(* IEC 61131-3 sources: labSCADA/project-view, 13 files *)

(* ---- FB_AnalogAlarm.st ---- *)
(* ==============================================================================
   FUNCTION BLOCK: FB_AnalogAlarm
   DESCRIPTION: IEC 61131-3 Structured Text implementation of an SEL RTAC-style
                analog alarm monitor with pickup/dropout hysteresis deadbands
                and sustained excursion / reset timers.

                Supports:
                - High Alarm trip / dropout (e.g. Fridge High > 8.0°C, reset < 7.5°C)
                - Low Alarm trip / dropout (e.g. Fridge Low < 2.0°C, reset > 2.5°C)
                - Window Alarm (High + Low simultaneously enabled)
                - Configurable Pickup Delay (prevents trips on brief door opens or noise)
                - Configurable Dropout Delay (anti-chatter filter on recovery)
                - Diagnostic Trip Outputs (HighTrip, LowTrip, Elapsed Timers)
   ============================================================================== *)
FUNCTION_BLOCK FB_AnalogAlarm
VAR_INPUT
	rVal            : REAL;             (* Analog process value to monitor (e.g. Temperature) *)
    bEnableHigh     : BOOL := TRUE;     (* Enable High Alarm monitoring *)
    rHighPickup     : REAL := 0.0;      (* High trip pickup threshold *)
    rHighDropout    : REAL := 0.0;      (* High trip reset threshold (or leave 0.0 and use rHysteresis) *)
    bEnableLow      : BOOL := FALSE;    (* Enable Low Alarm monitoring *)
    rLowPickup      : REAL := 0.0;      (* Low trip pickup threshold *)
    rLowDropout     : REAL := 0.0;      (* Low trip reset threshold (or leave 0.0 and use rHysteresis) *)
    rHysteresis     : REAL := 0.0;      (* Optional deadband offset applied if Dropout not explicitly set *)
    tPickupDelay    : TIME := T#0S;     (* Time excursion must persist before alarm asserts *)
    tDropoutDelay   : TIME := T#0S;     (* Time normal state must persist before alarm clears *)
END_VAR
VAR_OUTPUT
	bAlarm          : BOOL := FALSE;    (* Filtered alarm output (Active Alarm) *)
    bWarn           : BOOL := FALSE;    (* Pre-alarm warning: In excursion (pickup), timing towards alarm *)
    bPickup         : BOOL := FALSE;    (* Instantaneous pickup status (pre-timer) *)
    bHighTrip       : BOOL := FALSE;    (* TRUE if High Alarm condition caused/maintains trip *)
    bLowTrip        : BOOL := FALSE;    (* TRUE if Low Alarm condition caused/maintains trip *)
    tElapsedPU      : TIME := T#0S;     (* Current elapsed pickup timer *)
    tElapsedDO      : TIME := T#0S;     (* Current elapsed dropout timer *)
END_VAR
VAR
	rEffHighDO      : REAL;
    rEffLowDO       : REAL;
    bHighCondition  : BOOL := FALSE;
    bLowCondition   : BOOL := FALSE;
    fbTimer         : FB_PickupDropout;
END_VAR
// --- implementation ---
// 1. Calculate effective dropout thresholds
IF rHighDropout <> 0.0 THEN
    rEffHighDO := rHighDropout;
ELSIF rHysteresis > 0.0 THEN
    rEffHighDO := rHighPickup - rHysteresis;
ELSE
    rEffHighDO := rHighPickup;
END_IF;

IF rLowDropout <> 0.0 THEN
    rEffLowDO := rLowDropout;
ELSIF rHysteresis > 0.0 THEN
    rEffLowDO := rLowPickup + rHysteresis;
ELSE
    rEffLowDO := rLowPickup;
END_IF;

// 2. High threshold hysteresis evaluation
IF bEnableHigh THEN
    IF rVal >= rHighPickup THEN
        bHighCondition := TRUE;
    ELSIF rVal <= rEffHighDO THEN
        bHighCondition := FALSE;
    END_IF;
ELSE
    bHighCondition := FALSE;
END_IF;

// 3. Low threshold hysteresis evaluation
IF bEnableLow THEN
    IF rVal <= rLowPickup THEN
        bLowCondition := TRUE;
    ELSIF rVal >= rEffLowDO THEN
        bLowCondition := FALSE;
    END_IF;
ELSE
    bLowCondition := FALSE;
END_IF;

// 4. Pickup / Dropout timing filter (SEL RTAC PU_DO equivalent)
fbTimer(
    IN := (bHighCondition OR bLowCondition),
    tPickupDelay := tPickupDelay,
    tDropoutDelay := tDropoutDelay
);

bAlarm     := fbTimer.Q;
bPickup    := fbTimer.bPickup;
bWarn      := fbTimer.bPickup AND NOT fbTimer.Q;
tElapsedPU := fbTimer.tElapsedPU;
tElapsedDO := fbTimer.tElapsedDO;

// 5. Diagnostic cause flags
IF bAlarm THEN
    bHighTrip := bHighCondition;
    bLowTrip  := bLowCondition;
ELSE
    bHighTrip := FALSE;
    bLowTrip  := FALSE;
END_IF;
END_FUNCTION

(* ---- FB_APC_SmartUPS.st ---- *)
(* ==============================================================================
   FUNCTION BLOCK: FB_APC_SmartUPS
   DESCRIPTION: Encapsulated clinical monitoring block for UPS Power Systems
                following the Schneider Electric / APC Smart-UPS Modbus Register Map
                (AN-176 / 990-9840).
                - Supervised Utility Grid Power Loss (Generator Dispatch)
                - Battery State of Charge & Remaining Runtime Monitoring
                - Low Battery Reserve Emergency Escalation
                - Beeper Mute / Silence Supervisory Command Control
   ============================================================================== *)
FUNCTION_BLOCK FB_APC_SmartUPS
VAR_INPUT
    wStatusWord         : WORD := 16#0001;  (* Register 40001: Bit 0=Online, Bit 1=On Battery, Bit 4=Low Battery *)
    wBatteryPct         : WORD := 100;     (* Register 40002: Battery Charge (0-100%) *)
    wRuntimeSec         : WORD := 0;       (* Register 40003: Runtime in seconds *)
    wLineVoltageX10     : WORD := 1200;    (* Register 40004: Line Voltage * 10 (1200 = 120.0 V) *)
    wLoadPct            : WORD := 0;       (* Register 40005: Inverter Load (0-100%) *)
    wRuntimeMin         : WORD := 60;      (* Register 40007: Runtime in minutes *)
    wBeeperStatus       : WORD := 1;       (* Register 40008: 1=Enabled, 2=Muted, 3=Disabled *)

    (* --- Interactive Operator Commands (from Kiosk UI or PLC) --- *)
    bCmdMuteBeeper      : BOOL := FALSE;   (* TRUE pulse: Temporarily mute beeper for current power loss *)
    bCmdDisableBeeper   : BOOL := FALSE;   (* TRUE pulse: Disable beeper speaker *)
    bCmdEnableBeeper    : BOOL := FALSE;   (* TRUE pulse: Enable beeper speaker *)

    tPowerLossDelay     : TIME := T#10S;   (* Debounce filter to ignore momentary utility grid flickers *)
    wLowBatteryLimit    : WORD := 20;      (* Low battery alarm threshold (%) *)
    wLowRuntimeLimitMin : WORD := 15;      (* Low runtime alarm threshold (minutes) *)
END_VAR
VAR_OUTPUT
    bOnline             : BOOL := TRUE;    (* TRUE = Grid utility power is normal *)
    bOnBattery          : BOOL := FALSE;   (* TRUE = Running on battery inverter *)
    bAlarmPowerLost     : BOOL := FALSE;   (* Priority 2: Utility grid dropped -> Manual generator required *)
    bAlarmLowBattery    : BOOL := FALSE;   (* Priority 1: Battery reserve critically low *)
    rBatteryPct         : REAL := 100.0;   (* Battery % (0.0 - 100.0) *)
    rLineVoltage        : REAL := 120.0;   (* Utility line voltage in Volts RMS *)
    rRuntimeMinutes     : REAL := 60.0;    (* Estimated remaining runtime in minutes *)
    rLoadPct            : REAL := 0.0;     (* Current load percentage *)
    bBeeperMuted        : BOOL := FALSE;   (* Beeper is currently muted *)
    bBeeperDisabled     : BOOL := FALSE;   (* Beeper is disabled *)

    (* --- Modbus Command Output (Mapped to Holding Register 40010 / Offset 9) --- *)
    wCommandOut         : WORD := 0;       (* 1=Mute, 2=Disable, 3=Enable *)
END_VAR
VAR
    fbFilterPowerLoss   : FB_PickupDropout;
    tonCmdPulse         : TON;
    wActiveCmd          : WORD := 0;
    bPrevMute           : BOOL := FALSE;
    bPrevDisable        : BOOL := FALSE;
    bPrevEnable         : BOOL := FALSE;
END_VAR
// --- implementation ---
// 1. DECODE APC SMART-UPS STATUS WORD (Register 40001)
// Bit 0 = State Online (Grid OK)
// Bit 1 = State On Battery (Power Failure)
// Bit 4 = Low Battery
bOnline    := (wStatusWord AND 16#0001) <> 0;
bOnBattery := (wStatusWord AND 16#0002) <> 0;

// 2. CONVERT RAW TELEMETRY TO ENGINEERING UNITS
rBatteryPct     := WORD_TO_REAL(wBatteryPct);
rLineVoltage    := WORD_TO_REAL(wLineVoltageX10) / 10.0;
rLoadPct        := WORD_TO_REAL(wLoadPct);

// Beeper status
bBeeperMuted    := (wBeeperStatus = 2);
bBeeperDisabled := (wBeeperStatus = 3);

// Calculate runtime in minutes (prefer wRuntimeMin if non-zero, else wRuntimeSec / 60)
IF wRuntimeMin > 0 THEN
    rRuntimeMinutes := WORD_TO_REAL(wRuntimeMin);
ELSIF wRuntimeSec > 0 THEN
    rRuntimeMinutes := WORD_TO_REAL(wRuntimeSec) / 60.0;
ELSE
    rRuntimeMinutes := 0.0;
END_IF;

// 3. DEBOUNCED UTILITY POWER LOSS ALARM (Generator Dispatch)
// Ignores 1-2 second lightning flickers, trips after sustained outage (tPowerLossDelay)
fbFilterPowerLoss(
    IN            := bOnBattery,
    tPickupDelay  := tPowerLossDelay,
    tDropoutDelay := T#5S
);
bAlarmPowerLost := fbFilterPowerLoss.Q;

// 4. CRITICAL LOW BATTERY ALARM
// Triggers if battery % drops below limit OR runtime drops below critical threshold while on battery
IF bOnBattery AND ((wBatteryPct <= wLowBatteryLimit) OR (rRuntimeMinutes <= WORD_TO_REAL(wLowRuntimeLimitMin))) THEN
    bAlarmLowBattery := TRUE;
ELSE
    bAlarmLowBattery := FALSE;
END_IF;

// 5. BEEPER COMMAND EXECUTION (Pulsed Output to Modbus Register 40010)
// Latch active command for 1.5s so asynchronous Modbus cyclic task reliably transmits write
IF bCmdMuteBeeper AND NOT bPrevMute THEN
    wActiveCmd := 1;       // 1 = Mute
    bCmdMuteBeeper := FALSE;
ELSIF bCmdDisableBeeper AND NOT bPrevDisable THEN
    wActiveCmd := 2;       // 2 = Disable
    bCmdDisableBeeper := FALSE;
ELSIF bCmdEnableBeeper AND NOT bPrevEnable THEN
    wActiveCmd := 3;       // 3 = Enable
    bCmdEnableBeeper := FALSE;
END_IF;

bPrevMute    := bCmdMuteBeeper;
bPrevDisable := bCmdDisableBeeper;
bPrevEnable  := bCmdEnableBeeper;

tonCmdPulse(IN := (wActiveCmd > 0), PT := T#1500MS);
IF tonCmdPulse.Q THEN
    wActiveCmd := 0;
END_IF;

wCommandOut := wActiveCmd;
END_FUNCTION

(* ---- FB_Dewar.st ---- *)
(* ==============================================================================
   FUNCTION BLOCK: FB_Dewar
   DESCRIPTION: Encapsulated clinical monitoring block for Liquid Nitrogen (LN2)
                cryogenic storage vessels (dewars / freezers).
                - Scaled raw integer input (iRawTempX10 / 10.0 -> °C)
                - High threshold alarm with hysteresis & debounced pickup timing
                - Clinical fault supervision (Open circuit, wiring short, comms loss)
                - High-temperature excursion alarm gated off during hardware faults
                - Wireless cleanroom health diagnostics (Battery, RSSI, Watchdog, Faults)
   ============================================================================== *)
FUNCTION_BLOCK FB_Dewar
VAR_INPUT
    (* --- Operational Alarm Thresholds & Delays --- *)
    rHighTrip           : REAL := -135.0;   (* Critical specimen danger limit (°C) *)
    rHysteresis         : REAL := 5.0;      (* Reset deadband (°C) *)
    tPickupDelay        : TIME := T#30S;    (* Sustained warm excursion required to trip *)
    tDropoutDelay       : TIME := T#10S;    (* Clean fill required to reset *)

    (* --- 8 Modbus Holding Registers (Direct from Bridge Slot 1) --- *)
    wRawTempX10         : WORD := 16#D8F0;  (* Offset 0: Dewar scaled temp * 10 (-1954 = -195.4 °C, -9999 = Sentinel) *)
    uiRawBatteryMv      : UINT := 3850;     (* Offset 1: Battery health in millivolts *)
    uiRawFaultCode      : UINT := 0;        (* Offset 2: Probe fault (0=OK, 1=Open, 2=GND, 3=VCC, 4=Hardware Error) *)
    wRawRSSI            : WORD := 16#FFCE;  (* Offset 3: Wireless link margin in dBm (-50 = 16#FFCE) *)
    wRawSeqLow          : WORD := 0;        (* Offset 4: Sequence counter low word *)
    wRawSeqHigh         : WORD := 0;        (* Offset 5: Sequence counter high word *)
    uiRawAgeSec         : UINT := 0;        (* Offset 6: Telemetry age in seconds *)
    wRawStatusFlags     : WORD := 16#0001;  (* Offset 7: Bit 0=Online, Bit 1=LowBatt, Bit 2=CommLoss, Bit 3=AccessMode *)
    bIsWireless         : BOOL := TRUE;     (* TRUE = Enable wireless diagnostics *)
    tCommLossTimeout    : TIME := T#60S;    (* Watchdog comms loss alarm threshold *)

    (* --- Interactive Operator Commands (from Kiosk UI or OPC UA) --- *)
    bCmdSetAccessMode   : BOOL := FALSE;    (* TRUE pulse: Activate Access Mode (Alarms paused 30 min) *)
    bCmdCancelAccessMode: BOOL := FALSE;    (* TRUE pulse: Cancel Access Mode immediately *)
    rCalOffset          : REAL := 0.0;      (* NIST calibration trim offset in °C (clamped +/-10.0) *)
END_VAR
VAR_OUTPUT
    rProcessTemp        : REAL := -999.0;   (* Published process temperature to SCADA (°C) *)
    bAlarm              : BOOL := FALSE;    (* Priority 2 Emergency Temperature Alarm flag *)
    bWarn               : BOOL := FALSE;    (* Pre-alarm pickup delay warning flag *)
    rBatteryVolts       : REAL := 3.85;     (* Published battery voltage (V) *)
    bLowBattery         : BOOL := FALSE;    (* Low battery warning flag (< 3.4V) *)
    iRSSI               : INT := -50;       (* Published wireless link margin (dBm) *)
    bCommLoss           : BOOL := FALSE;    (* Comms loss watchdog alarm *)
    bProbeFault         : BOOL := TRUE;     (* Physical probe disconnected or shorted (defaults TRUE on cold boot) *)
    uiFaultCode         : UINT := 0;        (* Published probe fault reason (0=OK, 1=Open, 2=GND, 3=VCC) *)
    uiAgeSec            : UINT := 0;        (* Telemetry age in seconds *)
    bAccessMode         : BOOL := FALSE;    (* Access Mode active - Alarms paused 30 min for tank maintenance *)

    (* --- Modbus Command Outputs (Mapped to Bridge Holding Regs 10 & 11) --- *)
    wCommandMailboxOut  : WORD := 0;        (* Offset 10: 5 = SetAccessMode *)
    wCommandParamOut    : WORD := 0;        (* Offset 11: 30 = 30 minutes, 0 = Cancel *)
END_VAR
VAR
    iTempX10            : INT;
    fbAlarmEval         : FB_AnalogAlarm;
    wActiveCmdCode      : WORD := 0;
    wActiveCmdParam     : WORD := 0;
    bPrevSetAccess      : BOOL := FALSE;
    bPrevCancelAccess   : BOOL := FALSE;
    tonCmdPulse         : TON;
    rCalOffsetEff       : REAL := 0.0;
END_VAR
VAR CONSTANT
    cMaxCalOffset       : REAL := 10.0;
END_VAR
// --- implementation ---
// ==============================================================================
// 1. HARDWARE HEALTH & TELEMETRY DECODING
// ==============================================================================
// Explicitly cast Modbus unsigned WORD inputs to signed two's complement INT
iTempX10 := TO_INT(wRawTempX10);

IF bIsWireless THEN
    rBatteryVolts := TO_REAL(uiRawBatteryMv) / 1000.0;
    bLowBattery   := (uiRawBatteryMv < 3400) OR (wRawStatusFlags.1);
    iRSSI         := TO_INT(wRawRSSI);
    uiAgeSec      := uiRawAgeSec;
    uiFaultCode   := uiRawFaultCode;

    // Probe fault if hardware reported fault code or value is sentinel (<= -273°C or >= 900°C)
    bProbeFault   := (uiRawFaultCode <> 0) OR (iTempX10 <= -2730) OR (iTempX10 >= 9000);

    // Watchdog comms loss if bridge flagged or age exceeds timeout
    bCommLoss     := (NOT wRawStatusFlags.0) OR (wRawStatusFlags.2) OR (uiRawAgeSec > (TIME_TO_UINT(tCommLossTimeout) / 1000));

    // Access Mode Active (Bit 3 of status flags: Alarms paused 30 min)
    bAccessMode   := wRawStatusFlags.3;
ELSE
    rBatteryVolts := 0.0;
    bLowBattery   := FALSE;
    iRSSI         := 0;
    bCommLoss     := FALSE;
    uiFaultCode   := 0;
    bProbeFault   := (iTempX10 <= -2730) OR (iTempX10 >= 9000);
    uiAgeSec      := 0;
    bAccessMode   := FALSE;
END_IF;

// ==============================================================================
// 2. TEMPERATURE SENTINEL MAPPING
// ==============================================================================
IF rCalOffset > cMaxCalOffset THEN
    rCalOffsetEff := cMaxCalOffset;
ELSIF rCalOffset < -cMaxCalOffset THEN
    rCalOffsetEff := -cMaxCalOffset;
ELSE
    rCalOffsetEff := rCalOffset;
END_IF;

// If probe is faulted or comms lost, output standard invalid sentinel (-999.0 °C)
IF bProbeFault OR bCommLoss THEN
    rProcessTemp := -999.0;
ELSE
    rProcessTemp := (TO_REAL(iTempX10) / 10.0) + rCalOffsetEff;
END_IF;

// ==============================================================================
// 3. CLINICAL ALARM EVALUATION (Pickup / Dropout & Hysteresis)
// ==============================================================================
// Thermal excursion alarms are only evaluated when sensor data is valid and not in access mode
fbAlarmEval(
    rVal          := rProcessTemp,
    bEnableHigh   := NOT (bProbeFault OR bCommLoss OR bAccessMode),
    rHighPickup   := rHighTrip,
    rHighDropout  := rHighTrip - rHysteresis,
    bEnableLow    := FALSE,
    tPickupDelay  := tPickupDelay,
    tDropoutDelay := tDropoutDelay
);

// If in Access Mode, clamp alarms and warnings to FALSE immediately (bypassing dropout timer)
IF bAccessMode THEN
    bAlarm := FALSE;
    bWarn  := FALSE;
ELSE
    bAlarm := fbAlarmEval.bAlarm;
    bWarn  := fbAlarmEval.bWarn;
END_IF;

// ==============================================================================
// 4. SUPERVISORY COMMAND DISPATCH (Downlink to Bridge & Physical Node)
// ==============================================================================
// Latch active command for 2.0s so Modbus cyclic write task reliably transmits to Bridge
IF bCmdSetAccessMode AND NOT bPrevSetAccess THEN
    wActiveCmdCode    := 5;     // 5 = SetAccessMode
    wActiveCmdParam   := 30;    // 30 minutes
    bCmdSetAccessMode := FALSE;
ELSIF bCmdCancelAccessMode AND NOT bPrevCancelAccess THEN
    wActiveCmdCode       := 5;  // 5 = SetAccessMode
    wActiveCmdParam      := 0;  // 0 = Cancel / Normal Mode
    bCmdCancelAccessMode := FALSE;
END_IF;

bPrevSetAccess    := bCmdSetAccessMode;
bPrevCancelAccess := bCmdCancelAccessMode;

tonCmdPulse(IN := (wActiveCmdCode > 0), PT := T#2000MS);
IF tonCmdPulse.Q THEN
    wActiveCmdCode  := 0;
    wActiveCmdParam := 0;
END_IF;

wCommandMailboxOut := wActiveCmdCode;
wCommandParamOut   := wActiveCmdParam;
END_FUNCTION

(* ---- FB_FacilityDoor.st ---- *)
(* ==============================================================================
   FUNCTION BLOCK: FB_FacilityDoor
   DESCRIPTION: Encapsulated monitoring block for cleanroom and facility access doors
                (Main Entry, Procedure Room, Cryo Storage, Air Shower, Gown In/Out).
                Features:
                - Fail-safe normally closed contact supervision (24V/TRUE = Closed, 0V/FALSE = Open / Unwired)
                - Sustained open timer with contact chatter dropout filter (FB_PickupDropout)
                - Direct physical terminal binding (bDoorClosed)
                - Filtered alarm output to SCADA (bDoorAlarm)
   ============================================================================== *)
FUNCTION_BLOCK FB_FacilityDoor
VAR_INPUT
    bDoorClosed         : BOOL := FALSE;    (* Hardware DI: 24V/TRUE = Closed, 0V/FALSE = Open / Unwired *)
    tOpenAlarmDelay     : TIME := T#60M;    (* Sustained open threshold before alarm asserts *)
    tDropoutDelay       : TIME := T#5S;     (* Anti-chatter filter on door closure *)
END_VAR
VAR_OUTPUT
    bDoorAlarm          : BOOL := FALSE;    (* Filtered Priority 2 Alarm output to SCADA *)
END_VAR
VAR
    fbFilter            : FB_PickupDropout;
END_VAR
// --- implementation ---
// TIMED DEBOUNCE FILTER FOR DOOR HELD OPEN ALARM
fbFilter(
    IN            := NOT bDoorClosed,
    tPickupDelay  := tOpenAlarmDelay,
    tDropoutDelay := tDropoutDelay
);
bDoorAlarm := fbFilter.Q;
END_FUNCTION

(* ---- FB_G210_Incubator.st ---- *)
(* ==============================================================================
   FUNCTION BLOCK: FB_G210_Incubator
   DESCRIPTION: Encapsulated clinical monitoring block for K-Systems G210
                Multi-Chamber Incubators (10 Heated Zones).
                - 10 Chamber Zone Temperatures (Default -99.0°C unassigned sentinel)
                - Direct Physical Dry Alarm Contact (bAlarmContact)
                - Door/Recovery Mute Supervision (bMute)
                - Pickup/Dropout Debounce Filter
   ============================================================================== *)
FUNCTION_BLOCK FB_G210_Incubator
VAR_INPUT
    bAlarmContact       : BOOL := FALSE;    (* Physical dry alarm contact from incubator (Fail-Safe NC: TRUE = Normal/Closed, FALSE = Alarm/Open) *)
    bMute               : BOOL := FALSE;    (* TRUE = Suppress alarm (Cabinet door open or recovery grace) *)
    tPickupDelay        : TIME := T#15S;    (* Contact bounce filter *)
    tDropoutDelay       : TIME := T#5S;     (* Recovery confirmation filter *)
END_VAR
VAR_OUTPUT
    bAlarm              : BOOL := FALSE;    (* Filtered Priority 2 Alarm output to SCADA *)
    bMuted              : BOOL := FALSE;    (* Contact is tripped but actively suppressed by cabinet mute *)
    rZoneTemps          : ARRAY[1..10] OF REAL := [10(-99.0)];  (* 10 Heated Chambers, Default -99.0 °C (Unwired Sentinel) *)
END_VAR
VAR
    fbFilter            : FB_PickupDropout;
END_VAR
// --- implementation ---
// 1. TIMED DEBOUNCE FILTER ON FAIL-SAFE NC ALARM CONTACT (TRUE = Closed/Normal, FALSE = Open/Alarm)
fbFilter(
    IN            := NOT bAlarmContact,
    tPickupDelay  := tPickupDelay,
    tDropoutDelay := tDropoutDelay
);

// 2. MUTE SUPERVISION
// When bMute is TRUE (cabinet door open or grace period), suppress bAlarm.
bMuted := bMute AND fbFilter.Q;

IF bMute THEN
    bAlarm := FALSE;
ELSE
    bAlarm := fbFilter.Q;
END_IF;
END_FUNCTION

(* ---- FB_Incubator.st ---- *)
(* ==============================================================================
   FUNCTION BLOCK: FB_Incubator
   DESCRIPTION: Encapsulated clinical monitoring block for Embryology Incubators
                (benchtop trigas, box incubators) via discrete dry alarm contacts.
                Features:
                - Pickup/Dropout debounce filter (FB_PickupDropout)
                - Direct physical terminal binding (bAlarmContact)
                - Cabinet door / post-close mute supervision (bMute)
   ============================================================================== *)
FUNCTION_BLOCK FB_Incubator
VAR_INPUT
    bAlarmContact       : BOOL := FALSE;    (* Physical dry alarm contact from incubator (FALSE = Normal, TRUE = Alarm) *)
    bMute               : BOOL := FALSE;    (* TRUE = Suppress alarm (Cabinet door open or recovery grace) *)
    tPickupDelay        : TIME := T#15S;    (* Contact bounce suppression filter *)
    tDropoutDelay       : TIME := T#5S;     (* Recovery confirmation filter *)
END_VAR
VAR_OUTPUT
    bAlarm              : BOOL := FALSE;    (* Filtered Priority 2 Alarm output to SCADA *)
    bMuted              : BOOL := FALSE;    (* Contact is tripped but suppressed by active mute *)
END_VAR
VAR
    fbFilter            : FB_PickupDropout;
END_VAR
// --- implementation ---
// 1. TIMED DEBOUNCE FILTER
fbFilter(
    IN            := bAlarmContact,
    tPickupDelay  := tPickupDelay,
    tDropoutDelay := tDropoutDelay
);

// 2. MUTE SUPERVISION
// When bMute is active (cabinet door open or post-close grace), suppress bAlarm.
bMuted := bMute AND fbFilter.Q;

IF bMute THEN
    bAlarm := FALSE;
ELSE
    bAlarm := fbFilter.Q;
END_IF;
END_FUNCTION

(* ---- FB_IncubatorCabinet.st ---- *)
(* ==============================================================================
   FUNCTION BLOCK: FB_IncubatorCabinet
   DESCRIPTION: Enclosure microclimate and access supervision for benchtop
                incubator cabinet.
                Features:
                - Standardized fail-safe door contact supervision (Closed loop = Closed, Open loop = Open)
                - Autonomous incubator alarm muting while door is open
                - Post-closure recovery grace timer (TOF) to prevent nuisance alarms
                - Cabinet door left open alarm (TON)
                - Thermostatic exhaust fan control loop (hysteresis)
   ============================================================================== *)
FUNCTION_BLOCK FB_IncubatorCabinet
VAR_INPUT
    bDoorClosed         : BOOL := FALSE;    (* Hardware DI: 24V/TRUE = Closed, 0V/FALSE = Open / Disconnected *)
    tDoorAlarmDelay     : TIME := T#3M;     (* Alarm if cabinet door left open longer than this *)
    tPostCloseGrace     : TIME := T#3M;     (* Time to keep incubator alarms muted after door closes *)
    wRawTempX10         : WORD := 16#D8F0;  (* Raw Modbus 750-461 register x10 (244 = 24.4°C, -9999 = 16#D8F0) *)
    rFanOnSetpoint      : REAL := 28.0;     (* Exhaust fan ON setpoint in °C *)
    rFanHysteresis      : REAL := 1.5;      (* Deadband in °C (turns off at 26.5°C) *)
    rCalOffset          : REAL := 0.0;      (* NIST calibration trim offset in °C (clamped +/-10.0) *)
END_VAR
VAR_OUTPUT
    bDoorAlarm          : BOOL := FALSE;    (* Alarm: Cabinet door held open past delay *)
    bIncubatorMute      : BOOL := FALSE;    (* TRUE while door is open OR during post-closure grace *)
    tGraceRemaining     : TIME := T#0S;     (* Time remaining in post-close recovery grace *)
    bFanCommand         : BOOL := FALSE;    (* Command to future DO fan relay *)
    bCabinetOvertemp    : BOOL := FALSE;    (* Alarm: Cabinet internal temp >= 32°C *)
    rProcessTemp        : REAL := -999.0;   (* Published cabinet temperature (°C) to SCADA & DB *)
    bProbeFault         : BOOL := TRUE;     (* Physical RTD probe open/short/out-of-range fault *)
END_VAR
VAR
    tonDoorOpen         : TON;              (* Timer for door held open alert *)
    tofGrace            : TOF;              (* Off-delay timer keeping mute active post-closure *)
    iTempX10            : INT;
    rCalOffsetEff       : REAL := 0.0;
END_VAR
VAR CONSTANT
    cMaxCalOffset       : REAL := 10.0;
END_VAR
// --- implementation ---
// ==============================================================================
// 1. CABINET DOOR HELD OPEN ALARM
//    Fail-safe hardware: 24V (TRUE) when closed, 0V (FALSE) when open/cut.
// ==============================================================================
tonDoorOpen(
    IN := NOT bDoorClosed,
    PT := tDoorAlarmDelay
);
bDoorAlarm := tonDoorOpen.Q;

// ==============================================================================
// 2. INCUBATOR ALARM MUTING & POST-CLOSE RECOVERY GRACE (TOF)
// ==============================================================================
// While bDoorClosed is FALSE (door open), tofGrace.Q is TRUE.
// When bDoorClosed transitions to TRUE, tofGrace.Q STAYS TRUE for tPostCloseGrace.
tofGrace(
    IN := NOT bDoorClosed,
    PT := tPostCloseGrace
);
bIncubatorMute := tofGrace.Q;

// Compute remaining grace time while door is closed but timer is still running
IF bDoorClosed AND tofGrace.Q THEN
    tGraceRemaining := tPostCloseGrace - tofGrace.ET;
ELSE
    tGraceRemaining := T#0S;
END_IF;

// ==============================================================================
// 3. CABINET TEMPERATURE SCALING & PROBE FAULT SUPERVISION
// ==============================================================================
IF rCalOffset > cMaxCalOffset THEN
    rCalOffsetEff := cMaxCalOffset;
ELSIF rCalOffset < -cMaxCalOffset THEN
    rCalOffsetEff := -cMaxCalOffset;
ELSE
    rCalOffsetEff := rCalOffset;
END_IF;

iTempX10    := TO_INT(wRawTempX10);
bProbeFault := (iTempX10 <= -2000) OR (iTempX10 >= 8500);

IF bProbeFault THEN
    rProcessTemp := -999.0;
ELSE
    rProcessTemp := (TO_REAL(iTempX10) / 10.0) + rCalOffsetEff;
END_IF;

// ==============================================================================
// 4. THERMOSTATIC EXHAUST FAN CONTROL (HYSTERESIS)
// ==============================================================================
IF bProbeFault THEN
    bFanCommand := FALSE;
ELSIF rProcessTemp >= rFanOnSetpoint THEN
    bFanCommand := TRUE;
ELSIF rProcessTemp <= (rFanOnSetpoint - rFanHysteresis) THEN
    bFanCommand := FALSE;
END_IF;

// ==============================================================================
// 5. CABINET OVERTEMPERATURE SUPERVISION
// ==============================================================================
bCabinetOvertemp := (NOT bProbeFault) AND (rProcessTemp >= 32.0);
END_FUNCTION

(* ---- FB_MedColdStorage.st ---- *)
(* ==============================================================================
   FUNCTION BLOCK: FB_MedColdStorage
   DESCRIPTION: Encapsulated clinical monitoring block for Medical Cold Storage
                & Cleanroom Ambient Telemetry (Slot 2 Wireless Node).
                Integrates:
                - Medical Refrigerator (Hierarchical fbFridge: FB_MedFridge)
                - Medical Freezer (Hierarchical fbFreezer: FB_MedFreezer)
                - Lab Cleanroom Ambient Temp (20.0°C to 27.0°C Comfort Range)
                - Cleanroom Wireless Diagnostics (Battery, RSSI, Faults, Comm Loss)
                Modbus RTU Slave Slot 2 Holding Registers:
                - Offset 0: Mapped directly to fbFridge.wRawTempX10
                - Offsets 1..7: Shared wireless telemetry & diagnostics
                - Offset 8: Mapped directly to fbFreezer.wRawTempX10
                - Offset 9: Mapped to wRawAmbientTempX10
   ============================================================================== *)
FUNCTION_BLOCK FB_MedColdStorage
VAR_INPUT
    (* --- 10 Modbus Holding Registers (Direct from Bridge Slot 2) --- *)
    wRawFridgeTempX10   : WORD := 16#D8F0;  (* Offset 0: Raw Modbus register (Fridge scaled temp * 10, -9999 = 16#D8F0) *)
    uiRawBatteryMv      : UINT := 3820;     (* Offset 1: Battery health in millivolts *)
    uiRawFaultCode      : UINT := 0;        (* Offset 2: Probe fault code bitmask (bit 0=Fridge, bit 1=Freezer, bit 2=Ambient) *)
    wRawRSSI            : WORD := 16#FFCE;  (* Offset 3: Raw Modbus register (Link margin in dBm, -50 = 16#FFCE) *)
    wRawSeqLow          : WORD := 0;        (* Offset 4: Sequence counter low word *)
    wRawSeqHigh         : WORD := 0;        (* Offset 5: Sequence counter high word *)
    uiRawAgeSec         : UINT := 0;        (* Offset 6: Telemetry age in seconds *)
    wRawStatusFlags     : WORD := 16#0001;  (* Offset 7: Bit 0=Online, Bit 1=LowBatt, Bit 2=CommLoss *)
    wRawFreezerTempX10  : WORD := 16#D8F0;  (* Offset 8: Raw Modbus register (Freezer scaled temp * 10, -9999 = 16#D8F0) *)
    wRawAmbientTempX10  : WORD := 16#D8F0;  (* Offset 9: Raw Modbus register (Ambient scaled temp * 10, -9999 = 16#D8F0) *)

    (* --- Ambient Room Comfort Thresholds --- *)
    rAmbientHighTrip    : REAL := 27.0;     (* Cleanroom upper comfort limit (°C) *)
    rAmbientLowTrip     : REAL := 20.0;     (* Cleanroom lower comfort limit (°C) *)
    rAmbientHysteresis  : REAL := 0.5;      (* Anti-chatter deadband (°C) *)
    tAmbientPickupDelay : TIME := T#5M;     (* 5-minute sustained delay for HVAC drift *)
    tAmbientDropoutDelay: TIME := T#10S;    (* 10-second clean recovery *)

    bIsWireless         : BOOL := TRUE;     (* TRUE = Enable wireless diagnostics *)
    tCommLossTimeout    : TIME := T#60S;    (* Watchdog comms loss alarm threshold *)
    rAmbientCalOffset   : REAL := 0.0;      (* NIST calibration trim offset for Ambient °C (clamped +/-10.0) *)
END_VAR
VAR_OUTPUT
    (* --- Published Ambient Room Telemetry to SCADA & UI --- *)
    rAmbientTemp        : REAL := -999.0;   (* Cleanroom Ambient Room Temp (°C) *)
    bAmbientAlarm       : BOOL := FALSE;    (* Ambient Room Drift Priority 2 Alarm *)
    bAmbientWarn        : BOOL := FALSE;    (* Ambient Room Drift Warning *)
    bAmbientProbeFault  : BOOL := TRUE;     (* Ambient probe disconnected or shorted *)

    (* --- Shared Wireless Cleanroom Health Diagnostics --- *)
    rBatteryVolts       : REAL := 3.82;     (* Published battery voltage (V) *)
    bLowBattery         : BOOL := FALSE;    (* Low battery warning flag (< 3.4V) *)
    iRSSI               : INT := -50;       (* Published wireless link margin (dBm) *)
    bCommLoss           : BOOL := FALSE;    (* Comms loss watchdog alarm *)
    uiFaultCode         : UINT := 0;        (* Published probe fault reason *)
    uiAgeSec            : UINT := 0;        (* Telemetry age in seconds *)
END_VAR
VAR
    fbFridge            : FB_MedFridge;     (* Hierarchical Medical Refrigerator Subsystem *)
    fbFreezer           : FB_MedFreezer;    (* Hierarchical Medical Freezer Subsystem *)
    fbAmbientAlarmEval  : FB_AnalogAlarm;   (* Cleanroom Ambient Comfort Window Evaluator *)
    iAmbientTempX10     : INT;
    iFreezerTempX10     : INT;
    bFreezerSwapSuspect : BOOL := FALSE;
    uiFreezerFaultIn    : UINT := 0;
    rAmbCalOffsetEff    : REAL := 0.0;
    tonOnlineSettle     : TON;              (* Hold CommLoss through initial Modbus settle on boot/reconnect *)
    bLinkOnline         : BOOL := FALSE;    (* Bridge online bit set and watchdog healthy *)
END_VAR
VAR CONSTANT
    cMaxCalOffset       : REAL := 10.0;
END_VAR
// --- implementation ---
// ==============================================================================
// 1. SHARED WIRELESS CLEANROOM HEALTH & TELEMETRY DECODING
// ==============================================================================
IF bIsWireless THEN
    rBatteryVolts := TO_REAL(uiRawBatteryMv) / 1000.0;
    bLowBattery   := (uiRawBatteryMv < 3400) OR (wRawStatusFlags.1);
    iRSSI         := TO_INT(wRawRSSI);
    uiAgeSec      := uiRawAgeSec;
    uiFaultCode   := uiRawFaultCode;
    (* Require bridge Online bit (Bit 0) + 2s settle before leaving CommLoss
       so scan-1 unpopulated Modbus holding registers (all zeros = 0.0 C)
       cannot falsely prime the thermal vial filter on boot/reload. *)
    bLinkOnline   := wRawStatusFlags.0
        AND (NOT wRawStatusFlags.2)
        AND (uiRawAgeSec < (TIME_TO_UINT(tCommLossTimeout) / 1000));
    tonOnlineSettle(IN := bLinkOnline, PT := T#2S);
    bCommLoss     := NOT tonOnlineSettle.Q;
ELSE
    rBatteryVolts := 0.0;
    bLowBattery   := FALSE;
    iRSSI         := 0;
    bCommLoss     := FALSE;
    uiFaultCode   := 0;
    uiAgeSec      := 0;
    tonOnlineSettle(IN := FALSE);
END_IF;

// ==============================================================================
// 2. MEDICAL REFRIGERATOR (Hierarchical FB_MedFridge Instance)
// ==============================================================================
fbFridge(
    wRawTempX10         := wRawFridgeTempX10,
    uiRawFaultCode      := BOOL_TO_UINT((uiRawFaultCode AND 16#0001) <> 0),
    bCommLoss           := bCommLoss
);

// ==============================================================================
// 3. MEDICAL FREEZER (Hierarchical FB_MedFreezer Instance)
// ==============================================================================
(* Pre-evaluate Ambient fault & check for legacy dynamic-ROM slot shift
   (if Freezer probe drops out, pre-pinned node firmware shifts room Ambient
   >12 C into the Freezer slot while Ambient goes -999 / bit 2). *)
iAmbientTempX10     := TO_INT(wRawAmbientTempX10);
bAmbientProbeFault  := ((uiRawFaultCode AND 16#0004) <> 0) OR (iAmbientTempX10 <= -9000) OR (iAmbientTempX10 >= 9000);
iFreezerTempX10     := TO_INT(wRawFreezerTempX10);
bFreezerSwapSuspect := bAmbientProbeFault AND (iFreezerTempX10 > 120) AND (iFreezerTempX10 < 9000) AND (fbFreezer.rProcessTemp < 5.0);
uiFreezerFaultIn    := BOOL_TO_UINT(((uiRawFaultCode AND 16#0002) <> 0) OR bFreezerSwapSuspect);

fbFreezer(
    wRawTempX10         := wRawFreezerTempX10,
    uiRawFaultCode      := uiFreezerFaultIn,
    bCommLoss           := bCommLoss
);

// ==============================================================================
// 4. CLEANROOM AMBIENT ROOM TEMPERATURE (20.0°C to 27.0°C Comfort Window)
// ==============================================================================
IF rAmbientCalOffset > cMaxCalOffset THEN
    rAmbCalOffsetEff := cMaxCalOffset;
ELSIF rAmbientCalOffset < -cMaxCalOffset THEN
    rAmbCalOffsetEff := -cMaxCalOffset;
ELSE
    rAmbCalOffsetEff := rAmbientCalOffset;
END_IF;

IF bAmbientProbeFault OR bCommLoss THEN
    rAmbientTemp := -999.0;
ELSE
    rAmbientTemp := (TO_REAL(iAmbientTempX10) / 10.0) + rAmbCalOffsetEff;
END_IF;

fbAmbientAlarmEval(
    rVal          := rAmbientTemp,
    bEnableHigh   := NOT (bAmbientProbeFault OR bCommLoss),
    rHighPickup   := rAmbientHighTrip,
    rHighDropout  := rAmbientHighTrip - rAmbientHysteresis,
    bEnableLow    := NOT (bAmbientProbeFault OR bCommLoss),
    rLowPickup    := rAmbientLowTrip,
    rLowDropout   := rAmbientLowTrip + rAmbientHysteresis,
    tPickupDelay  := tAmbientPickupDelay,
    tDropoutDelay := tAmbientDropoutDelay
);
bAmbientAlarm := fbAmbientAlarmEval.bAlarm;
bAmbientWarn  := fbAmbientAlarmEval.bWarn;
END_FUNCTION

(* ---- FB_MedFreezer.st ---- *)
(* ==============================================================================
   FUNCTION BLOCK: FB_MedFreezer
   DESCRIPTION: Encapsulated clinical monitoring block for Medical Freezers
                (-20°C sperm/media or -80°C ultra-low freezers).
                - Scaled raw integer input (wRawTempX10 / 10.0 -> °C)
                - First-order thermal mass filter (FB_ThermalVial) emulating a buffer vial
                - High temperature threshold alarm on virtual-vial temperature
                - Option A pre-alarm warning (bWarn) from temperature margin band
                - Clinical fault supervision (Open circuit, wiring short, comms loss)
   ============================================================================== *)
FUNCTION_BLOCK FB_MedFreezer
VAR_INPUT
    wRawTempX10         : WORD := 16#D8F0;  (* Offset 0: Raw Modbus register (-9999 = 16#D8F0 Sentinel / Disconnected) *)
    rHighTrip           : REAL := -10.0;    (* Medications/consumables warm alarm threshold (°C) per USP <1079> *)
    rHysteresis         : REAL := 0.5;      (* Anti-chatter deadband (°C) - resets at -10.5°C *)
    tPickupDelay        : TIME := T#0S;     (* Binary pickup delay (T#0S when using virtual-vial damping) *)
    tDropoutDelay       : TIME := T#0S;     (* Binary dropout delay (hysteresis handles anti-chatter) *)
    tThermalTau         : TIME := T#8M;     (* Virtual buffer vial time constant; T#0S bypasses filtering *)
    rHighWarnMargin     : REAL := 2.0;      (* Pre-alarm warn margin below rHighTrip (-12.0°C when High=-10.0°C) *)
    uiRawFaultCode      : UINT := 0;        (* Probe fault code: 0=OK, 0xFF=Unpopulated *)
    bCommLoss           : BOOL := FALSE;    (* Watchdog comms loss flag *)
    rCalOffset          : REAL := 0.0;      (* NIST calibration trim offset in °C (clamped +/-10.0) *)
END_VAR
VAR_OUTPUT
    rProcessTemp        : REAL := -999.0;   (* Virtual-vial temperature to SCADA & DB (°C) *)
    rRawTemp            : REAL := -999.0;   (* Instantaneous unfiltered air temperature (°C) *)
    bAlarm              : BOOL := FALSE;    (* Priority 2 Emergency Alarm flag *)
    bWarn               : BOOL := FALSE;    (* Priority 1 Pre-alarm warning flag (margin band or pickup delay) *)
    bProbeFault         : BOOL := TRUE;     (* Probe disconnected or hardware fault *)
END_VAR
VAR
    iTempX10            : INT;
    bHealthy            : BOOL;
    bProcessValid       : BOOL;
    rCalOffsetEff       : REAL := 0.0;
    fbThermalVial       : FB_ThermalVial;
    fbAlarmEval         : FB_AnalogAlarm;
    fbWarnEval          : FB_AnalogAlarm;
END_VAR
VAR CONSTANT
    cMaxCalOffset       : REAL := 10.0;
END_VAR
// --- implementation ---
// ==============================================================================
// 1. HARDWARE HEALTH & RAW AIR TEMPERATURE SCALING
// ==============================================================================
IF rCalOffset > cMaxCalOffset THEN
    rCalOffsetEff := cMaxCalOffset;
ELSIF rCalOffset < -cMaxCalOffset THEN
    rCalOffsetEff := -cMaxCalOffset;
ELSE
    rCalOffsetEff := rCalOffset;
END_IF;

iTempX10    := TO_INT(wRawTempX10);
bProbeFault := (uiRawFaultCode <> 0) OR (iTempX10 <= -9000) OR (iTempX10 >= 9000);
bHealthy    := NOT (bProbeFault OR bCommLoss);

IF NOT bHealthy THEN
    rRawTemp := -999.0;
ELSE
    rRawTemp := (TO_REAL(iTempX10) / 10.0) + rCalOffsetEff;
END_IF;

// ==============================================================================
// 2. VIRTUAL BUFFER VIAL FILTER (8-Minute Thermal Time Constant)
// ==============================================================================
fbThermalVial(
    rRawTemp    := rRawTemp,
    bValid      := bHealthy,
    tThermalTau := tThermalTau,
    rCalOffset  := rCalOffsetEff
);
rProcessTemp := fbThermalVial.rVialTemp;
bProcessValid := (rProcessTemp > -273.0) AND (rProcessTemp < 900.0);

// ==============================================================================
// 3. CLINICAL ALARM & PRE-ALARM MARGIN EVALUATION
// ==============================================================================
fbAlarmEval(
    rVal          := rProcessTemp,
    bEnableHigh   := bProcessValid,
    rHighPickup   := rHighTrip,
    rHighDropout  := rHighTrip - rHysteresis,
    bEnableLow    := FALSE,
    rHysteresis   := rHysteresis,
    tPickupDelay  := tPickupDelay,
    tDropoutDelay := tDropoutDelay
);

fbWarnEval(
    rVal        := rProcessTemp,
    bEnableHigh := bProcessValid AND (rHighWarnMargin > 0.0),
    rHighPickup := rHighTrip - rHighWarnMargin,
    rHysteresis := rHysteresis,
    bEnableLow  := FALSE
);

bAlarm := fbAlarmEval.bAlarm;
bWarn  := fbAlarmEval.bWarn OR (fbWarnEval.bAlarm AND NOT fbAlarmEval.bAlarm);
END_FUNCTION

(* ---- FB_MedFridge.st ---- *)
(* ==============================================================================
   FUNCTION BLOCK: FB_MedFridge
   DESCRIPTION: Encapsulated clinical monitoring block for Medical Refrigerators
                (embryo media, medications, specimens).
                - Scaled raw integer input (wRawTempX10 / 10.0 -> °C)
                - First-order thermal mass filter (FB_ThermalVial) emulating a buffer vial
                - Dual-limit Window Alarm (1.0°C to 8.5°C/10.0°C) on virtual-vial temp
                - Option A pre-alarm warning (bWarn) from temperature margin bands
                - Clinical fault supervision (Open circuit, wiring short, comms loss)
   ============================================================================== *)
FUNCTION_BLOCK FB_MedFridge
VAR_INPUT
    wRawTempX10         : WORD := 16#D8F0;  (* Raw Modbus register (Fridge scaled temp * 10, -9999 = 16#D8F0) *)
    rHighTrip           : REAL := 8.5;      (* CAP excursion threshold (override to 10.0 in AFOA PLC_PRG) *)
    rLowTrip            : REAL := 1.0;      (* Freezing prevention threshold (1.0°C clinical alarm per equipment.json) *)
    rHysteresis         : REAL := 0.5;      (* Anti-chatter deadband (°C) *)
    tPickupDelay        : TIME := T#0S;     (* Binary pickup delay (T#0S when using virtual-vial damping) *)
    tDropoutDelay       : TIME := T#0S;     (* Binary dropout delay (hysteresis handles anti-chatter) *)
    tThermalTau         : TIME := T#5M;     (* Virtual buffer vial time constant; T#0S bypasses filtering *)
    rHighWarnMargin     : REAL := 1.5;      (* Pre-alarm warn margin below rHighTrip (8.5°C when High=10.0°C) *)
    rLowWarnMargin      : REAL := 1.0;      (* Pre-alarm warn margin above rLowTrip (2.0°C when Low=1.0°C) *)
    uiRawFaultCode      : UINT := 0;        (* Probe fault code: 0=OK, 0xFF=Unpopulated *)
    bCommLoss           : BOOL := FALSE;    (* Watchdog comms loss flag *)
    rCalOffset          : REAL := 0.0;      (* NIST calibration trim offset in °C (clamped +/-10.0) *)
END_VAR
VAR_OUTPUT
    rProcessTemp        : REAL := -999.0;   (* Virtual-vial temperature to SCADA & DB (°C) *)
    rRawTemp            : REAL := -999.0;   (* Instantaneous unfiltered air temperature (°C) *)
    bAlarm              : BOOL := FALSE;    (* Priority 2 Emergency Alarm flag *)
    bWarn               : BOOL := FALSE;    (* Priority 1 Pre-alarm warning flag (margin band or pickup delay) *)
    bProbeFault         : BOOL := TRUE;     (* Physical probe disconnected or shorted *)
END_VAR
VAR
    iTempX10            : INT;
    bHealthy            : BOOL;
    bProcessValid       : BOOL;
    rCalOffsetEff       : REAL := 0.0;
    fbThermalVial       : FB_ThermalVial;
    fbAlarmEval         : FB_AnalogAlarm;
    fbWarnEval          : FB_AnalogAlarm;
END_VAR
VAR CONSTANT
    cZero               : REAL := 0.0;
    cMaxCalOffset       : REAL := 10.0;
END_VAR
// --- implementation ---
// ==============================================================================
// 1. HARDWARE HEALTH & RAW AIR TEMPERATURE SCALING
// ==============================================================================
IF rCalOffset > cMaxCalOffset THEN
    rCalOffsetEff := cMaxCalOffset;
ELSIF rCalOffset < -cMaxCalOffset THEN
    rCalOffsetEff := -cMaxCalOffset;
ELSE
    rCalOffsetEff := rCalOffset;
END_IF;

iTempX10    := TO_INT(wRawTempX10);
bProbeFault := (uiRawFaultCode <> 0) OR (iTempX10 <= -9000) OR (iTempX10 >= 9000);
bHealthy    := NOT (bProbeFault OR bCommLoss);

IF NOT bHealthy THEN
    rRawTemp := -999.0;
ELSE
    rRawTemp := (TO_REAL(iTempX10) / 10.0) + rCalOffsetEff;
END_IF;

// ==============================================================================
// 2. VIRTUAL BUFFER VIAL FILTER (5-Minute Thermal Time Constant)
// ==============================================================================
fbThermalVial(
    rRawTemp    := rRawTemp,
    bValid      := bHealthy,
    tThermalTau := tThermalTau,
    rCalOffset  := rCalOffsetEff
);
rProcessTemp := fbThermalVial.rVialTemp;
bProcessValid := (rProcessTemp > -273.0) AND (rProcessTemp < 900.0);

// ==============================================================================
// 3. CLINICAL ALARM & PRE-ALARM MARGIN EVALUATION (Dual-Limit Window)
// ==============================================================================
fbAlarmEval(
    rVal          := rProcessTemp,
    bEnableHigh   := bProcessValid,
    rHighPickup   := rHighTrip,
    rHighDropout  := rHighTrip - rHysteresis,
    bEnableLow    := bProcessValid,
    rLowPickup    := rLowTrip,
    rLowDropout   := rLowTrip + rHysteresis,
    rHysteresis   := rHysteresis,
    tPickupDelay  := tPickupDelay,
    tDropoutDelay := tDropoutDelay
);

fbWarnEval(
    rVal        := rProcessTemp,
    bEnableHigh := bProcessValid AND (rHighWarnMargin > cZero),
    rHighPickup := rHighTrip - rHighWarnMargin,
    bEnableLow  := bProcessValid AND (rLowWarnMargin > cZero),
    rLowPickup  := rLowTrip + rLowWarnMargin,
    rHysteresis := rHysteresis
);

bAlarm := fbAlarmEval.bAlarm;
bWarn  := fbAlarmEval.bWarn OR (fbWarnEval.bAlarm AND NOT fbAlarmEval.bAlarm);
END_FUNCTION

(* ---- FB_PickupDropout.st ---- *)
(* ==============================================================================
   FUNCTION BLOCK: FB_PickupDropout
   DESCRIPTION: IEC 61131-3 Structured Text implementation of the SEL RTAC
                Pickup / Dropout timer (equivalent to RTAC PU_DO).

                - Pickup Delay (On-Delay / Timeout):
                  The input signal (IN) must remain continuously TRUE for
                  tPickupDelay before the output (Q) asserts to TRUE.
                  Nuisance spikes or transients shorter than tPickupDelay
                  are filtered out and reset the timer.

                - Dropout Delay (Off-Delay / Chatter Filter):
                  Once Q is TRUE (tripped), IN must remain continuously FALSE
                  for tDropoutDelay before Q resets to FALSE.
                  Any bounce or re-trip during the dropout window resets
                  the dropout timer, keeping Q asserted.
   ============================================================================== *)
FUNCTION_BLOCK FB_PickupDropout
VAR_INPUT
	IN              : BOOL;             (* Input signal to evaluate *)
    tPickupDelay    : TIME := T#0S;     (* Time IN must be sustained TRUE before Q asserts *)
    tDropoutDelay   : TIME := T#0S;     (* Time IN must be sustained FALSE before Q deasserts *)
END_VAR
VAR_OUTPUT
	Q               : BOOL := FALSE;    (* Filtered output state *)
    bPickup         : BOOL := FALSE;    (* Raw instantaneous input status (unfiltered) *)
    tElapsedPU      : TIME := T#0S;     (* Elapsed pickup timer *)
    tElapsedDO      : TIME := T#0S;     (* Elapsed dropout timer *)
END_VAR
VAR
	tonPickup       : TON;
    tonDropout      : TON;
END_VAR
// --- implementation ---
// Track raw instantaneous input
bPickup := IN;

IF NOT Q THEN
    // --- Alarm is currently OFF: Timing towards Pickup ---
    tonDropout(IN := FALSE, PT := tDropoutDelay);
    tElapsedDO := T#0S;

    tonPickup(IN := IN, PT := tPickupDelay);
    tElapsedPU := tonPickup.ET;

    IF tonPickup.Q THEN
        Q := TRUE;
    END_IF;
ELSE
    // --- Alarm is currently ON: Timing towards Dropout ---
    tonPickup(IN := FALSE, PT := tPickupDelay);
    tElapsedPU := tPickupDelay;

    tonDropout(IN := NOT IN, PT := tDropoutDelay);
    tElapsedDO := tonDropout.ET;

    IF tonDropout.Q THEN
        Q := FALSE;
    END_IF;
END_IF;
END_FUNCTION

(* ---- FB_RandomGenerator.st ---- *)
FUNCTION_BLOCK FB_RandomGenerator
VAR_INPUT
    bExecute: BOOL; (* Set TRUE to calculate next random number *)
    diMin: DINT; (* Inclusive minimum value *)
    diMax: DINT; (* Inclusive maximum value *)
END_VAR
VAR_OUTPUT
    diResult: DINT; (* Generated random number *)
END_VAR
VAR
    udiSeed: UDINT := 123456789; (* Initial non-zero seed *)
    udiRange: UDINT;
END_VAR
// --- implementation ---
IF bExecute THEN
    (* LCG Formula: X_{n+1} = (a * X_n + c) mod 2^32 *)
    udiSeed := (udiSeed * 1664525) + 1013904223;

    (* Scale the 32-bit value to the requested [diMin..diMax] range *)
    IF diMax >= diMin THEN
        udiRange := DINT_TO_UDINT(diMax - diMin + 1);
        diResult := diMin + UDINT_TO_DINT(udiSeed MOD udiRange);
    ELSE
        diResult := diMin;
    END_IF;
END_IF;
END_FUNCTION_BLOCK

(* ---- FB_ThermalVial.st ---- *)
(* ==============================================================================
   FUNCTION BLOCK: FB_ThermalVial
   DESCRIPTION: First-order thermal mass low-pass filter (EWMA) emulating a
                temperature sensor immersed in a glycol, mineral-oil, or sand vial.
                - Scan-rate independent discrete update driven by tSampleTick
                - Instant seed on cold boot or recovery from probe/comms fault
                - Hold last buffered value across transient probe/comms dropouts up to tHoldoverGrace
                - Revert to -999.0 only after holdover expires (or immediately if never primed)
                - Set tThermalTau := T#0S for zero-lag raw pass-through
   ============================================================================== *)
FUNCTION_BLOCK FB_ThermalVial
VAR_INPUT
    rRawTemp            : REAL := -999.0;   (* Instantaneous valid air temperature (°C) *)
    bValid              : BOOL := FALSE;    (* TRUE when probe & comms are healthy *)
    tThermalTau         : TIME := T#5M;     (* First-order thermal time constant tau; T#0S bypasses filter *)
    tSampleTick         : TIME := T#5S;     (* Fixed EWMA update interval dt *)
    tHoldoverGrace      : TIME := T#5M;     (* Max holdover across brief dropouts; T#0S disables holdover *)
    rCalOffset          : REAL := 0.0;      (* Upstream calibration trim; step changes shift primed filter state *)
END_VAR
VAR_OUTPUT
    rVialTemp           : REAL := -999.0;   (* Buffered virtual-vial temperature (°C), or -999.0 if invalid *)
END_VAR
VAR
    tonTick             : TON;
    tonHoldover         : TON;
    rFilteredTemp       : REAL := -999.0;
    bPrimed             : BOOL := FALSE;
    bInputOk            : BOOL := FALSE;
    tEffTick            : TIME;
    diDtMs              : DINT;
    diTauMs             : DINT;
    rAlpha              : REAL;
    rPrevCalOffset      : REAL := 0.0;
    bCalTrackInit       : BOOL := FALSE;
    rOffsetDelta        : REAL := 0.0;
END_VAR
VAR CONSTANT
    cTempInvalid        : REAL := -999.0;
    cTempMinValid       : REAL := -273.0;
    cTempMaxValid       : REAL := 900.0;
    cTimeZero           : TIME := T#0S;
    cDefaultSampleTick  : TIME := T#5S;
END_VAR
// --- implementation ---
IF NOT bCalTrackInit THEN
    rPrevCalOffset := rCalOffset;
    bCalTrackInit  := TRUE;
    rOffsetDelta   := 0.0;
ELSIF rCalOffset <> rPrevCalOffset THEN
    rOffsetDelta   := rCalOffset - rPrevCalOffset;
    rPrevCalOffset := rCalOffset;
ELSE
    rOffsetDelta   := 0.0;
END_IF;

bInputOk := bValid AND (rRawTemp > cTempMinValid) AND (rRawTemp < cTempMaxValid);
IF tSampleTick > cTimeZero THEN
    tEffTick := tSampleTick;
ELSE
    tEffTick := cDefaultSampleTick;
END_IF;

IF NOT bInputOk THEN
    tonTick(IN := FALSE, PT := tEffTick);
    IF bPrimed AND (tHoldoverGrace > cTimeZero) THEN
        tonHoldover(IN := TRUE, PT := tHoldoverGrace);
        IF tonHoldover.Q THEN
            tonHoldover(IN := FALSE, PT := tHoldoverGrace);
            bPrimed       := FALSE;
            rFilteredTemp := cTempInvalid;
        ELSIF rOffsetDelta <> 0.0 THEN
            rFilteredTemp := rFilteredTemp + rOffsetDelta;
        END_IF;
    ELSE
        tonHoldover(IN := FALSE, PT := tHoldoverGrace);
        bPrimed       := FALSE;
        rFilteredTemp := cTempInvalid;
    END_IF;
ELSIF (tThermalTau <= cTimeZero) OR (NOT bPrimed) THEN
    tonHoldover(IN := FALSE, PT := tHoldoverGrace);
    bPrimed       := TRUE;
    rFilteredTemp := rRawTemp;
    tonTick(IN := FALSE, PT := tEffTick);
ELSE
    IF rOffsetDelta <> 0.0 THEN
        rFilteredTemp := rFilteredTemp + rOffsetDelta;
    END_IF;
    tonHoldover(IN := FALSE, PT := tHoldoverGrace);
    tonTick(IN := TRUE, PT := tEffTick);
    IF tonTick.Q THEN
        tonTick(IN := FALSE, PT := tEffTick);
        diDtMs        := TIME_TO_DINT(tEffTick);
        diTauMs       := TIME_TO_DINT(tThermalTau);
        rAlpha        := TO_REAL(diDtMs) / TO_REAL(diTauMs + diDtMs);
        rFilteredTemp := rFilteredTemp + rAlpha * (rRawTemp - rFilteredTemp);
    END_IF;
END_IF;

rVialTemp := rFilteredTemp;
END_FUNCTION_BLOCK
